// TIA Portal V14 SP1 export
// export: Created 2000-01-01T00:00:00.0000000Z, ExportSetting None
DATA_BLOCK "MCP_RC_DB6"   // DB9806
{ S7_Optimized_Access := 'TRUE' }
   VAR
      Count : Int := 2;
      D : "MCP_RC_UDT3";
   END_VAR
BEGIN
END_DATA_BLOCK
